Fanuc KAREL source: KT00769.KL

PROGRAM KT00769
%NOLOCKGROUP
VAR
  B1: BOOLEAN
  B2: BOOLEAN
  OUT: REAL
BEGIN
  B1 = TRUE
  B2 = FALSE
  B1 = TRUE
  B2 = FALSE
  OUT = ACOS(B1)
END KT00769
